ABB RAPID module: PrecProg.mod

MODULE MainModule
GLOBAL VAR robtarget robpoint0= p:{{-640.585, 506.981, 371.534},{0.375352, 0.284211, 0.854623, -0.218985}}{cfg 0,-1,2,0}{EJ 0.000000000,0.000000000,0.000000000,0.000000000,0.000000000,0.000000000}
GLOBAL VAR robtarget robpoint1= p:{{0.500, -0.500, 0.250},{0.000000, 1.000000, 0.000044, 0.000044}}{cfg -1,0,-2,0}{EJ 0.000000000,0.000000000,0.000000000,0.000000000,0.000000000,0.000000000}
GLOBAL VAR robtarget robpoint2= p:{{1500.120, -2000.990, -10.500},{0.707107, -0.000000, 0.707107, -0.000000}}{cfg -1,0,-2,0}{EJ 0.000000000,0.000000000,0.000000000,0.000000000,0.000000000,0.000000000}
GLOBAL VAR robtarget robpoint3= p:{{-353.026, -90.135, 331.702},{0.344329, 0.048056, 0.933073, -0.092215}}{cfg 0,-1,2,0}{EJ 0.000000000,0.000000000,0.000000000,0.000000000,0.000000000,0.000000000}

GLOBAL Proc main()
    wobj16.x = 0.0004
    wobj16.y = -0.001
    wobj16.z = 1000.000
    wobj16.q1 = 0.707097
    wobj16.q2 = 0.707102
    wobj16.q3 = -0.002324
    wobj16.q4 = 0.003847
    tool03.x = 0.125
    tool03.y = -0.375
    tool03.z = 123.457
    tool03.q1 = 0.923042
    tool03.q2 = -0.384698
    tool03.q3 = -0.000000
    tool03.q4 = 0.000001
    MoveL robpoint0,v50,z50,tool03,wobj16
    MoveL robpoint1,v50,z50,tool03,wobj16
    MoveJ robpoint2,v50,z50,tool03,wobj16
    Wait 0.002
    Wait 1.000
    MoveL robpoint3,v66,z50,tool03,wobj16
EndProc
EndModule
